(* IEC 61131-3 sources: kns-pump-station/tests/POUs/Fakes/FB_FakeEventSink, 8 files *)

(* ---- FB_FakeEventSink.decl.st ---- *)
// Назначение: подменный журнал событий станции для юнит-тестов (I_StationEventSink): кольцо 16
//             последних событий (код и значение), счётчик всех событий, поиск по коду.
// Автор:      kr0nsch
// Версия:     0.1.0
// Документ:   docs/DESIGN.md, раздел 6.14
FUNCTION_BLOCK FB_FakeEventSink IMPLEMENTS I_StationEventSink
VAR CONSTANT
    RING_LAST : UINT := 15;         // кольцо 0…15: 16 последних событий
END_VAR
VAR_OUTPUT
    udiCount   : UDINT;             // событий с последнего Clear
    eLastEvent : E_StationEvent;    // последнее событие
    rLastValue : REAL;              // его значение
END_VAR
VAR
    aeRing : ARRAY[0..RING_LAST] OF E_StationEvent;   // коды событий
    arRing : ARRAY[0..RING_LAST] OF REAL;             // значения
    uiHead : UINT;                  // индекс следующей записи
END_VAR

(* ---- CountOf.method.decl.st ---- *)
// Сколько событий с кодом eFind среди последних 16
METHOD PUBLIC CountOf : UINT
VAR_INPUT
    eFind : E_StationEvent;         // искомый код
END_VAR
VAR
    uiIdx  : UINT;                  // элемент кольца
    uiUsed : UINT;                  // заполнено элементов
END_VAR

(* ---- CountOf.method.impl.st ---- *)
CountOf := 0;
IF udiCount > RING_LAST THEN
    uiUsed := RING_LAST + 1;
ELSE
    uiUsed := UDINT_TO_UINT(udiCount);
END_IF
FOR uiIdx := 0 TO RING_LAST DO
    IF uiIdx < uiUsed AND aeRing[uiIdx] = eFind THEN
        CountOf := CountOf + 1;
    END_IF
END_FOR

(* ---- Has.method.decl.st ---- *)
// Есть ли событие eFind среди последних 16
METHOD PUBLIC Has : BOOL
VAR_INPUT
    eFind : E_StationEvent;         // искомый код
END_VAR

(* ---- LogEvent.method.decl.st ---- *)
// Записать событие в кольцо (самое старое затирается); всегда TRUE
METHOD PUBLIC LogEvent : BOOL
VAR_INPUT
    eEvent : E_StationEvent;        // код события
    rValue : REAL;                  // значение
END_VAR

(* ---- LogEvent.method.impl.st ---- *)
aeRing[uiHead] := eEvent;
arRing[uiHead] := rValue;
IF uiHead >= RING_LAST THEN
    uiHead := 0;
ELSE
    uiHead := uiHead + 1;
END_IF
udiCount := udiCount + 1;
eLastEvent := eEvent;
rLastValue := rValue;
LogEvent := TRUE;

(* ---- ValueOf.method.decl.st ---- *)
// Значение самого нового события eFind среди последних 16; нет такого — -1
METHOD PUBLIC ValueOf : REAL
VAR_INPUT
    eFind : E_StationEvent;         // искомый код
END_VAR
VAR
    uiStep  : UINT;                 // шаг назад от новейшего
    uiIdx   : UINT;                 // элемент кольца
    xFound  : BOOL;                 // найдено
END_VAR

(* ---- ValueOf.method.impl.st ---- *)
ValueOf := -1.0;
xFound := FALSE;
uiIdx := uiHead;
FOR uiStep := 0 TO RING_LAST DO
    IF uiIdx = 0 THEN
        uiIdx := RING_LAST;
    ELSE
        uiIdx := uiIdx - 1;
    END_IF
    IF NOT xFound AND UINT_TO_UDINT(uiStep) < udiCount AND aeRing[uiIdx] = eFind THEN
        ValueOf := arRing[uiIdx];
        xFound := TRUE;
    END_IF
END_FOR
